// Mitsubishi GX Works2 project: B_v6_d23   PLC: Q03UDE

PROGRAM COMMON
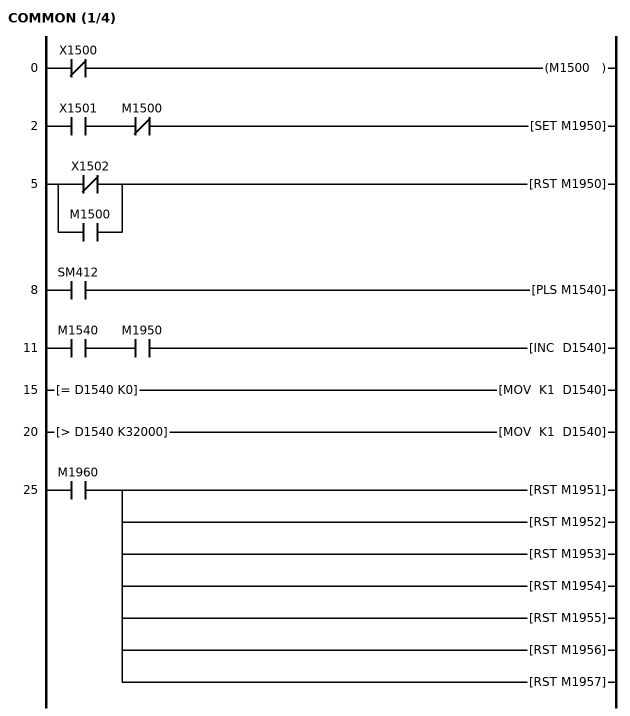
0     LDI     X1500
      OUT     M1500
2     LD      X1501
      ANI     M1500
      SET     M1950
5     LDI     X1502
      OR      M1500
      RST     M1950
8     LD      SM412
      PLS     M1540
11    LD      M1540
      AND     M1950
      INC     D1540
15    LD=     D1540 K0
      MOV     K1 D1540
20    LD>     D1540 K32000
      MOV     K1 D1540
25    LD      M1960
      RST     M1951
      RST     M1952
      RST     M1953
      RST     M1954
      RST     M1955
      RST     M1956
      RST     M1957
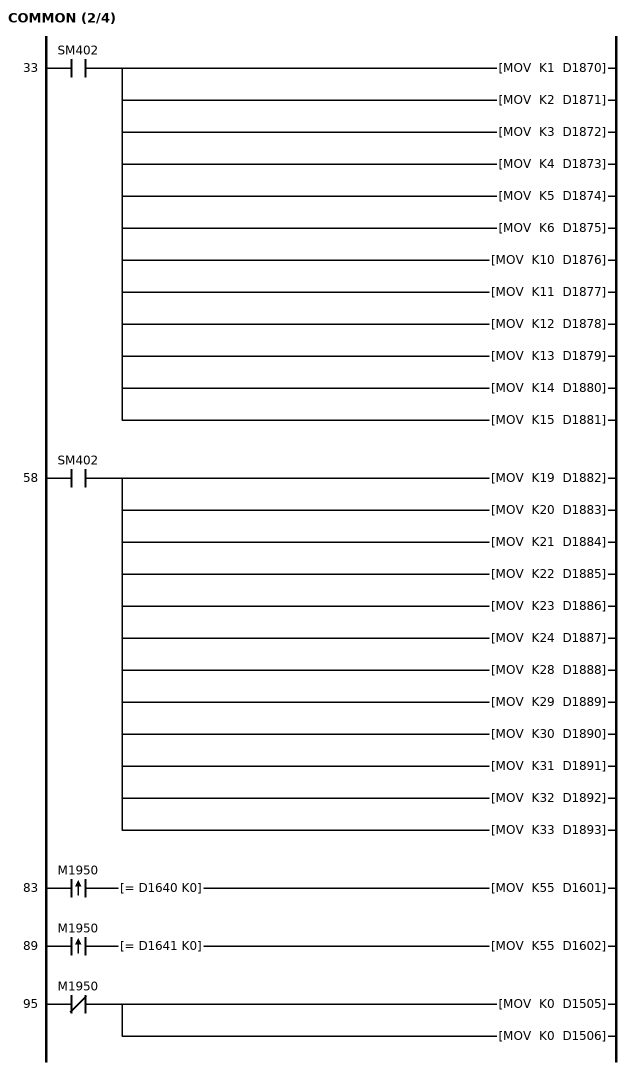
33    LD      SM402
      MOV     K1 D1870
      MOV     K2 D1871
      MOV     K3 D1872
      MOV     K4 D1873
      MOV     K5 D1874
      MOV     K6 D1875
      MOV     K10 D1876
      MOV     K11 D1877
      MOV     K12 D1878
      MOV     K13 D1879
      MOV     K14 D1880
      MOV     K15 D1881
58    LD      SM402
      MOV     K19 D1882
      MOV     K20 D1883
      MOV     K21 D1884
      MOV     K22 D1885
      MOV     K23 D1886
      MOV     K24 D1887
      MOV     K28 D1888
      MOV     K29 D1889
      MOV     K30 D1890
      MOV     K31 D1891
      MOV     K32 D1892
      MOV     K33 D1893
83    LDP     M1950
      AND=    D1640 K0
      MOV     K55 D1601
89    LDP     M1950
      AND=    D1641 K0
      MOV     K55 D1602
95    LDI     M1950
      MOV     K0 D1505
      MOV     K0 D1506
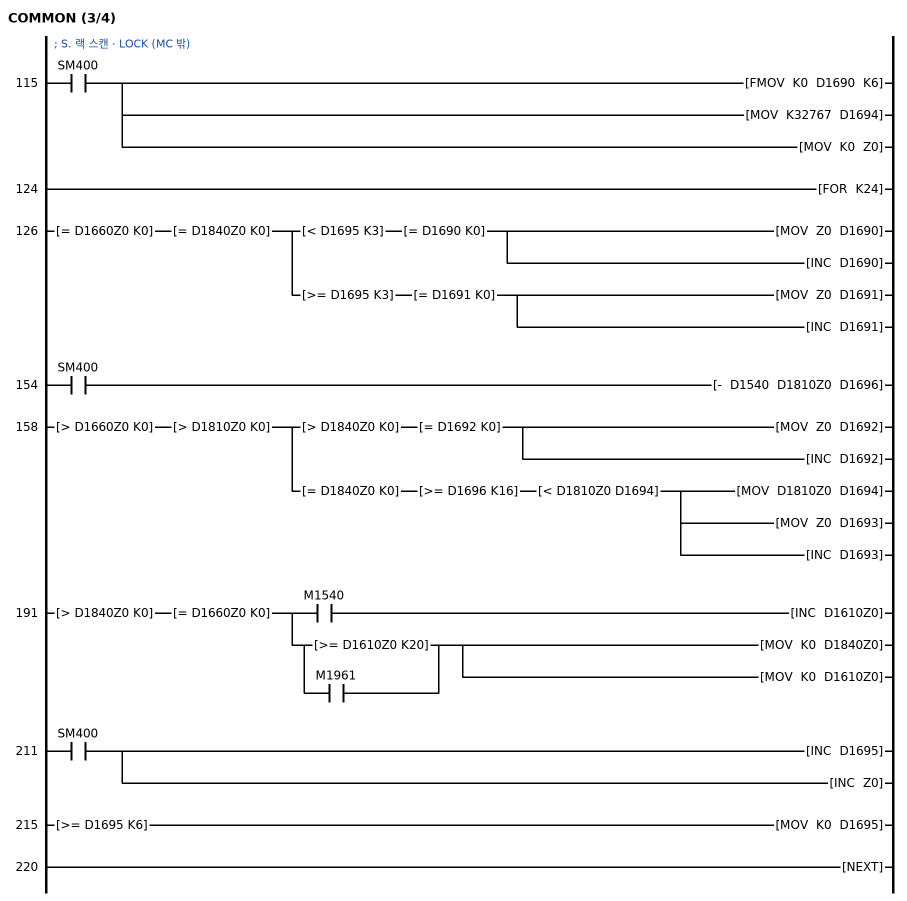
; S. 랙 스캔 · LOCK (MC 밖)
115   LD      SM400
      FMOV    K0 D1690 K6
      MOV     K32767 D1694
      MOV     K0 Z0
124   FOR     K24
126   LD=     D1660Z0 K0
      AND=    D1840Z0 K0
      MPS
      AND<    D1695 K3
      AND=    D1690 K0
      MOV     Z0 D1690
      INC     D1690
      MPP
      AND>=   D1695 K3
      AND=    D1691 K0
      MOV     Z0 D1691
      INC     D1691
154   LD      SM400
      -       D1540 D1810Z0 D1696
158   LD>     D1660Z0 K0
      AND>    D1810Z0 K0
      MPS
      AND>    D1840Z0 K0
      AND=    D1692 K0
      MOV     Z0 D1692
      INC     D1692
      MPP
      AND=    D1840Z0 K0
      AND>=   D1696 K16
      AND<    D1810Z0 D1694
      MOV     D1810Z0 D1694
      MOV     Z0 D1693
      INC     D1693
191   LD>     D1840Z0 K0
      AND=    D1660Z0 K0
      MPS
      AND     M1540
      INC     D1610Z0
      MPP
      LD>=    D1610Z0 K20
      OR      M1961
      ANB
      MOV     K0 D1840Z0
      MOV     K0 D1610Z0
211   LD      SM400
      INC     D1695
      INC     Z0
215   LD>=    D1695 K6
      MOV     K0 D1695
220   NEXT
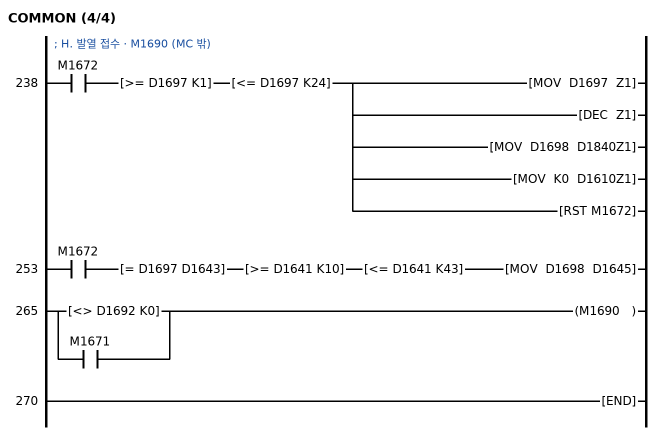
; H. 발열 접수 · M1690 (MC 밖)
238   LD      M1672
      AND>=   D1697 K1
      AND<=   D1697 K24
      MOV     D1697 Z1
      DEC     Z1
      MOV     D1698 D1840Z1
      MOV     K0 D1610Z1
      RST     M1672
253   LD      M1672
      AND=    D1697 D1643
      AND>=   D1641 K10
      AND<=   D1641 K43
      MOV     D1698 D1645
265   LD<>    D1692 K0
      OR      M1671
      OUT     M1690
270   END
END_PROGRAM

PROGRAM RFID
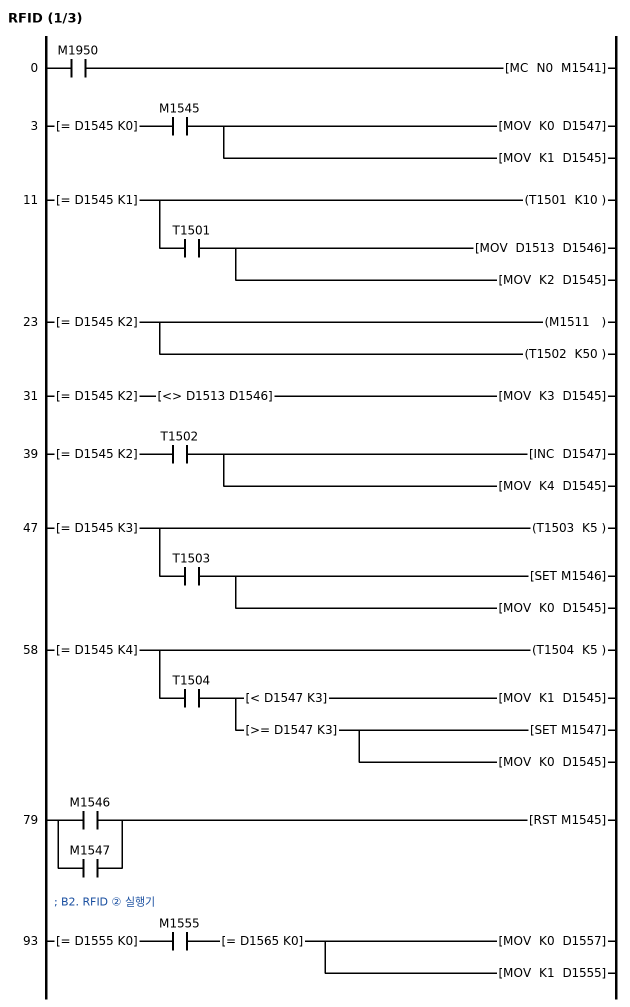
0     LD      M1950
      MC      N0 M1541
3     LD=     D1545 K0
      AND     M1545
      MOV     K0 D1547
      MOV     K1 D1545
11    LD=     D1545 K1
      OUT     T1501 K10
      AND     T1501
      MOV     D1513 D1546
      MOV     K2 D1545
23    LD=     D1545 K2
      OUT     M1511
      OUT     T1502 K50
31    LD=     D1545 K2
      AND<>   D1513 D1546
      MOV     K3 D1545
39    LD=     D1545 K2
      AND     T1502
      INC     D1547
      MOV     K4 D1545
47    LD=     D1545 K3
      OUT     T1503 K5
      AND     T1503
      SET     M1546
      MOV     K0 D1545
58    LD=     D1545 K4
      OUT     T1504 K5
      AND     T1504
      MPS
      AND<    D1547 K3
      MOV     K1 D1545
      MPP
      AND>=   D1547 K3
      SET     M1547
      MOV     K0 D1545
79    LD      M1546
      OR      M1547
      RST     M1545
; B2. RFID ② 실행기
93    LD=     D1555 K0
      AND     M1555
      AND=    D1565 K0
      MOV     K0 D1557
      MOV     K1 D1555
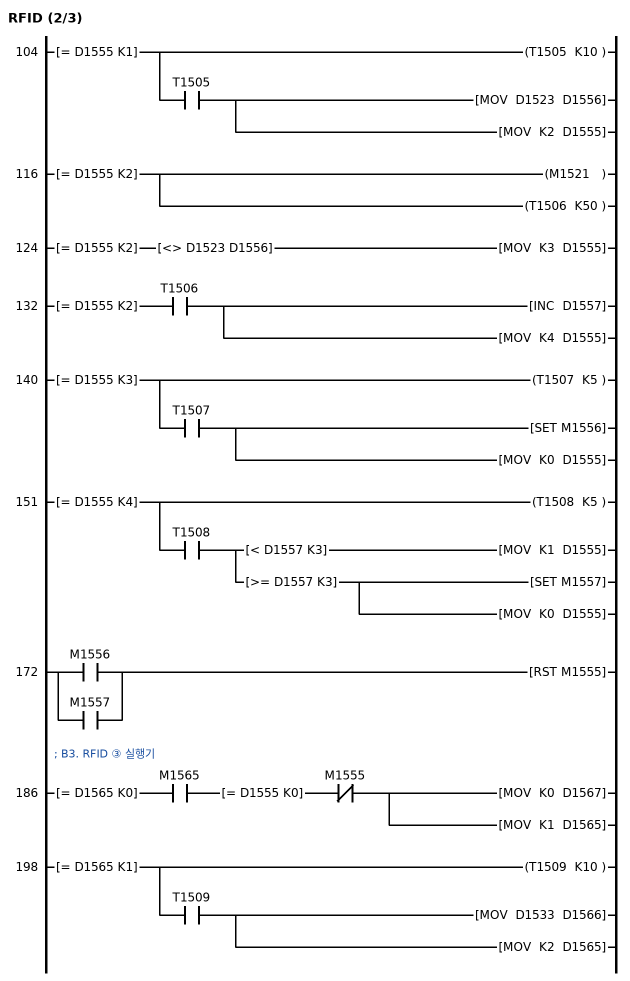
104   LD=     D1555 K1
      OUT     T1505 K10
      AND     T1505
      MOV     D1523 D1556
      MOV     K2 D1555
116   LD=     D1555 K2
      OUT     M1521
      OUT     T1506 K50
124   LD=     D1555 K2
      AND<>   D1523 D1556
      MOV     K3 D1555
132   LD=     D1555 K2
      AND     T1506
      INC     D1557
      MOV     K4 D1555
140   LD=     D1555 K3
      OUT     T1507 K5
      AND     T1507
      SET     M1556
      MOV     K0 D1555
151   LD=     D1555 K4
      OUT     T1508 K5
      AND     T1508
      MPS
      AND<    D1557 K3
      MOV     K1 D1555
      MPP
      AND>=   D1557 K3
      SET     M1557
      MOV     K0 D1555
172   LD      M1556
      OR      M1557
      RST     M1555
; B3. RFID ③ 실행기
186   LD=     D1565 K0
      AND     M1565
      AND=    D1555 K0
      ANI     M1555
      MOV     K0 D1567
      MOV     K1 D1565
198   LD=     D1565 K1
      OUT     T1509 K10
      AND     T1509
      MOV     D1533 D1566
      MOV     K2 D1565
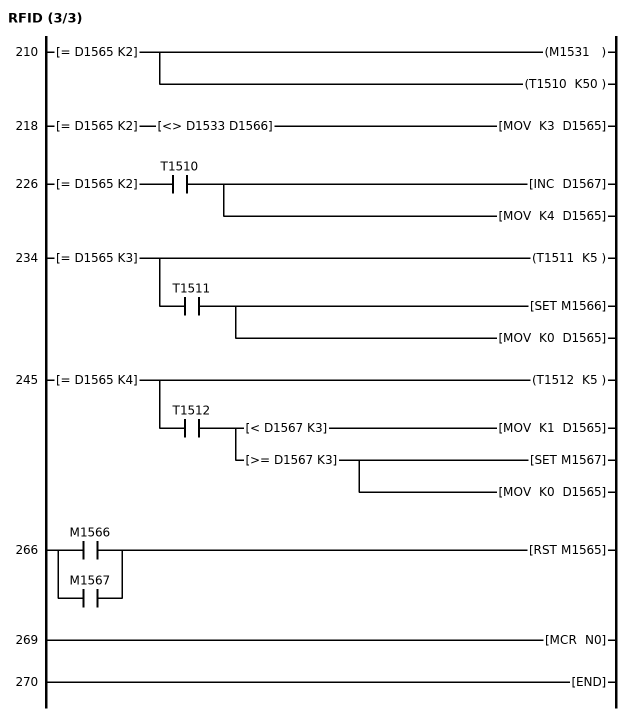
210   LD=     D1565 K2
      OUT     M1531
      OUT     T1510 K50
218   LD=     D1565 K2
      AND<>   D1533 D1566
      MOV     K3 D1565
226   LD=     D1565 K2
      AND     T1510
      INC     D1567
      MOV     K4 D1565
234   LD=     D1565 K3
      OUT     T1511 K5
      AND     T1511
      SET     M1566
      MOV     K0 D1565
245   LD=     D1565 K4
      OUT     T1512 K5
      AND     T1512
      MPS
      AND<    D1567 K3
      MOV     K1 D1565
      MPP
      AND>=   D1567 K3
      SET     M1567
      MOV     K0 D1565
266   LD      M1566
      OR      M1567
      RST     M1565
269   MCR     N0
270   END
END_PROGRAM

PROGRAM INFEED
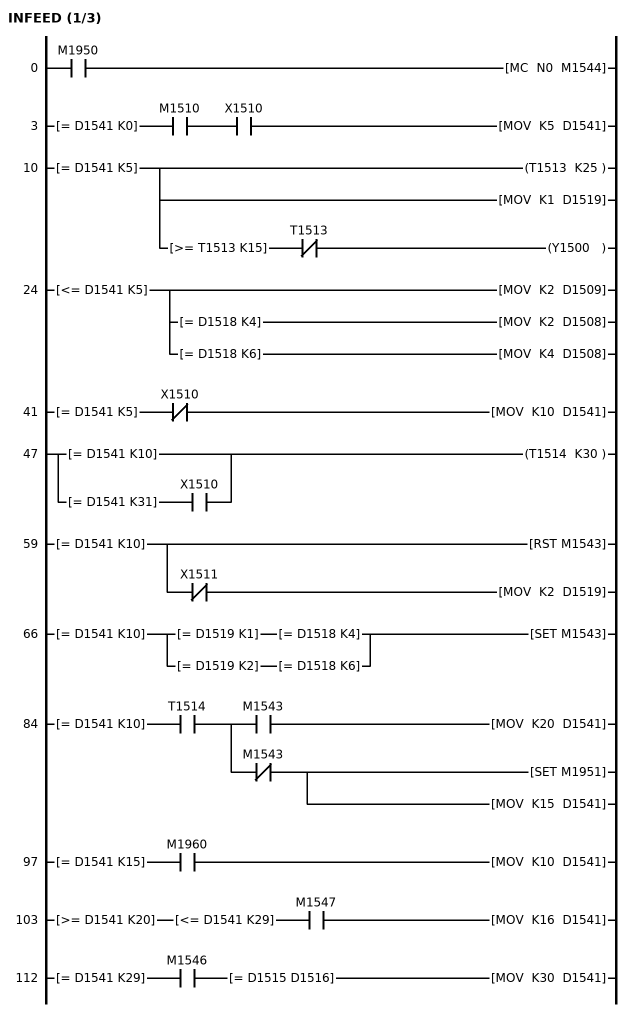
0     LD      M1950
      MC      N0 M1544
3     LD=     D1541 K0
      AND     M1510
      AND     X1510
      MOV     K5 D1541
10    LD=     D1541 K5
      OUT     T1513 K25
      MOV     K1 D1519
      AND>=   T1513 K15
      ANI     T1513
      OUT     Y1500
24    LD<=    D1541 K5
      MOV     K2 D1509
      MPS
      AND=    D1518 K4
      MOV     K2 D1508
      MPP
      AND=    D1518 K6
      MOV     K4 D1508
41    LD=     D1541 K5
      ANI     X1510
      MOV     K10 D1541
47    LD=     D1541 K10
      LD=     D1541 K31
      AND     X1510
      ORB
      OUT     T1514 K30
59    LD=     D1541 K10
      RST     M1543
      ANI     X1511
      MOV     K2 D1519
66    LD=     D1541 K10
      LD=     D1519 K1
      AND=    D1518 K4
      LD=     D1519 K2
      AND=    D1518 K6
      ORB
      ANB
      SET     M1543
84    LD=     D1541 K10
      AND     T1514
      MPS
      AND     M1543
      MOV     K20 D1541
      MPP
      ANI     M1543
      SET     M1951
      MOV     K15 D1541
97    LD=     D1541 K15
      AND     M1960
      MOV     K10 D1541
103   LD>=    D1541 K20
      AND<=   D1541 K29
      AND     M1547
      MOV     K16 D1541
112   LD=     D1541 K29
      AND     M1546
      AND=    D1515 D1516
      MOV     K30 D1541
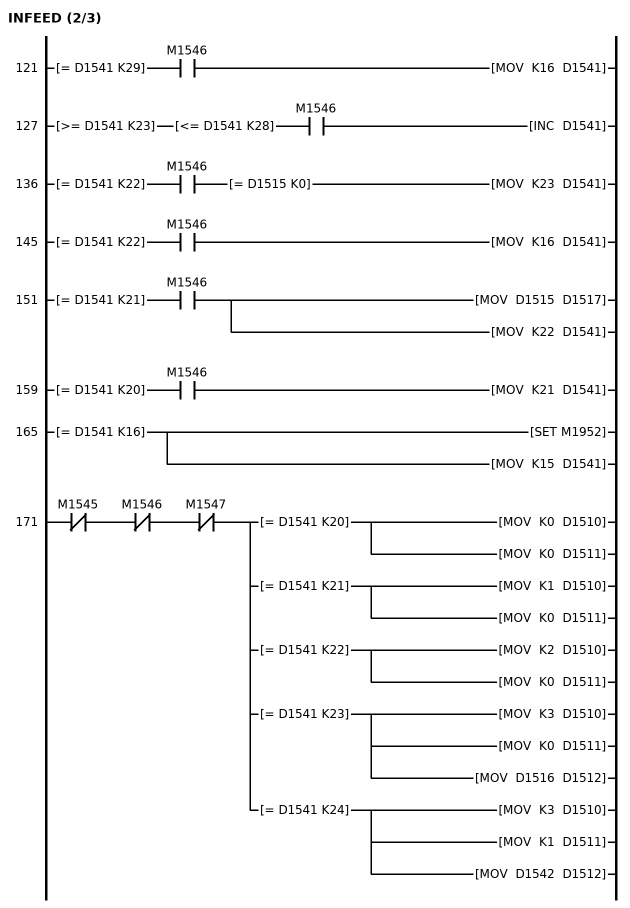
121   LD=     D1541 K29
      AND     M1546
      MOV     K16 D1541
127   LD>=    D1541 K23
      AND<=   D1541 K28
      AND     M1546
      INC     D1541
136   LD=     D1541 K22
      AND     M1546
      AND=    D1515 K0
      MOV     K23 D1541
145   LD=     D1541 K22
      AND     M1546
      MOV     K16 D1541
151   LD=     D1541 K21
      AND     M1546
      MOV     D1515 D1517
      MOV     K22 D1541
159   LD=     D1541 K20
      AND     M1546
      MOV     K21 D1541
165   LD=     D1541 K16
      SET     M1952
      MOV     K15 D1541
171   LDI     M1545
      ANI     M1546
      ANI     M1547
      MPS
      AND=    D1541 K20
      MOV     K0 D1510
      MOV     K0 D1511
      MRD
      AND=    D1541 K21
      MOV     K1 D1510
      MOV     K0 D1511
      MRD
      AND=    D1541 K22
      MOV     K2 D1510
      MOV     K0 D1511
      MRD
      AND=    D1541 K23
      MOV     K3 D1510
      MOV     K0 D1511
      MOV     D1516 D1512
      MPP
      AND=    D1541 K24
      MOV     K3 D1510
      MOV     K1 D1511
      MOV     D1542 D1512
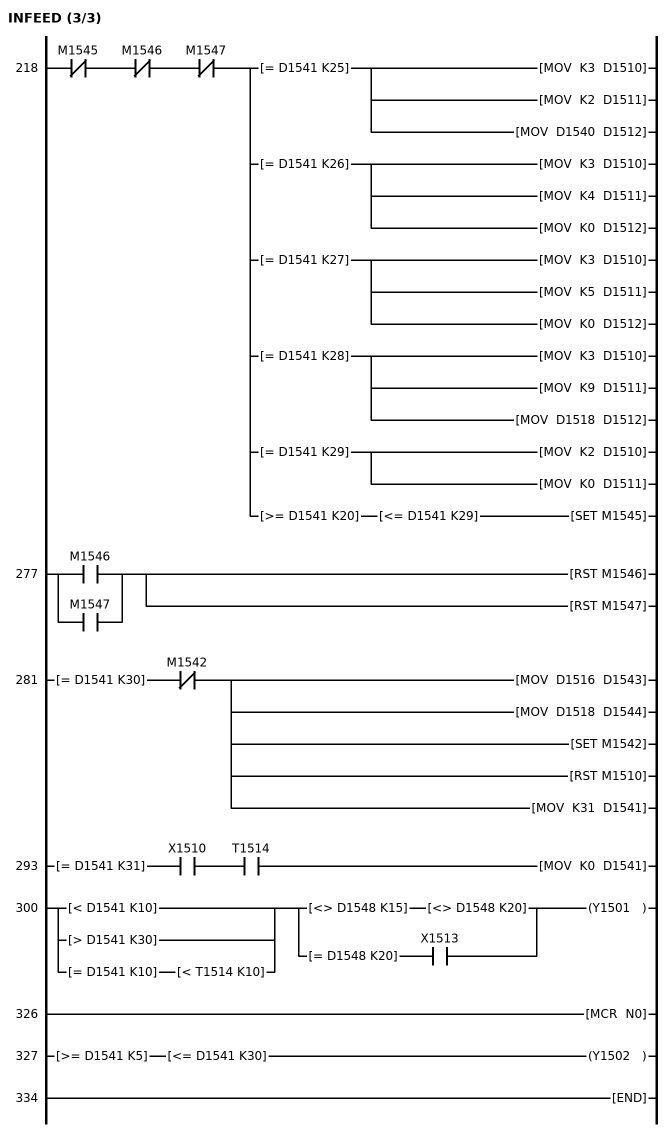
218   LDI     M1545
      ANI     M1546
      ANI     M1547
      MPS
      AND=    D1541 K25
      MOV     K3 D1510
      MOV     K2 D1511
      MOV     D1540 D1512
      MRD
      AND=    D1541 K26
      MOV     K3 D1510
      MOV     K4 D1511
      MOV     K0 D1512
      MRD
      AND=    D1541 K27
      MOV     K3 D1510
      MOV     K5 D1511
      MOV     K0 D1512
      MRD
      AND=    D1541 K28
      MOV     K3 D1510
      MOV     K9 D1511
      MOV     D1518 D1512
      MRD
      AND=    D1541 K29
      MOV     K2 D1510
      MOV     K0 D1511
      MPP
      AND>=   D1541 K20
      AND<=   D1541 K29
      SET     M1545
277   LD      M1546
      OR      M1547
      RST     M1546
      RST     M1547
281   LD=     D1541 K30
      ANI     M1542
      MOV     D1516 D1543
      MOV     D1518 D1544
      SET     M1542
      RST     M1510
      MOV     K31 D1541
293   LD=     D1541 K31
      AND     X1510
      AND     T1514
      MOV     K0 D1541
300   LD<     D1541 K10
      OR>     D1541 K30
      LD=     D1541 K10
      AND<    T1514 K10
      ORB
      LD<>    D1548 K15
      AND<>   D1548 K20
      LD=     D1548 K20
      AND     X1513
      ORB
      ANB
      OUT     Y1501
326   MCR     N0
327   LD>=    D1541 K5
      AND<=   D1541 K30
      OUT     Y1502
334   END
END_PROGRAM

PROGRAM CRANE
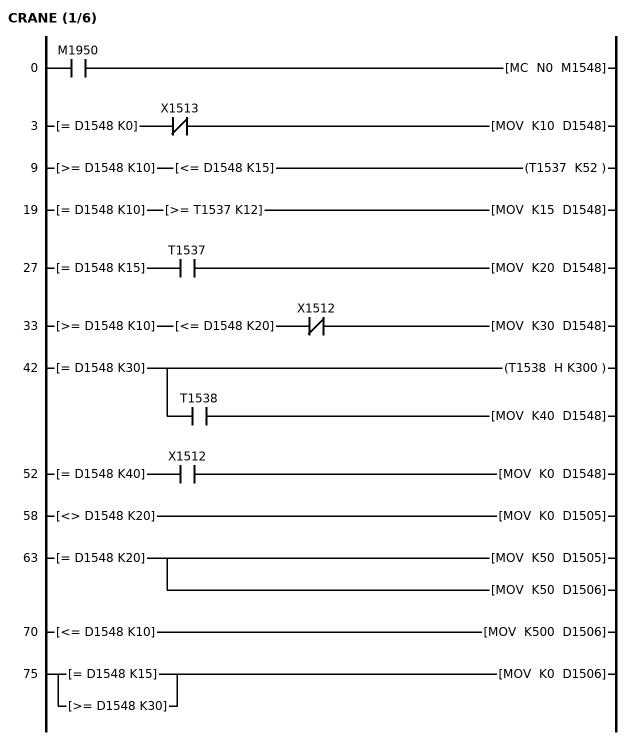
0     LD      M1950
      MC      N0 M1548
3     LD=     D1548 K0
      ANI     X1513
      MOV     K10 D1548
9     LD>=    D1548 K10
      AND<=   D1548 K15
      OUT     T1537 K52
19    LD=     D1548 K10
      AND>=   T1537 K12
      MOV     K15 D1548
27    LD=     D1548 K15
      AND     T1537
      MOV     K20 D1548
33    LD>=    D1548 K10
      AND<=   D1548 K20
      ANI     X1512
      MOV     K30 D1548
42    LD=     D1548 K30
      OUTH    T1538 K300
      AND     T1538
      MOV     K40 D1548
52    LD=     D1548 K40
      AND     X1512
      MOV     K0 D1548
58    LD<>    D1548 K20
      MOV     K0 D1505
63    LD=     D1548 K20
      MOV     K50 D1505
      MOV     K50 D1506
70    LD<=    D1548 K10
      MOV     K500 D1506
75    LD=     D1548 K15
      OR>=    D1548 K30
      MOV     K0 D1506
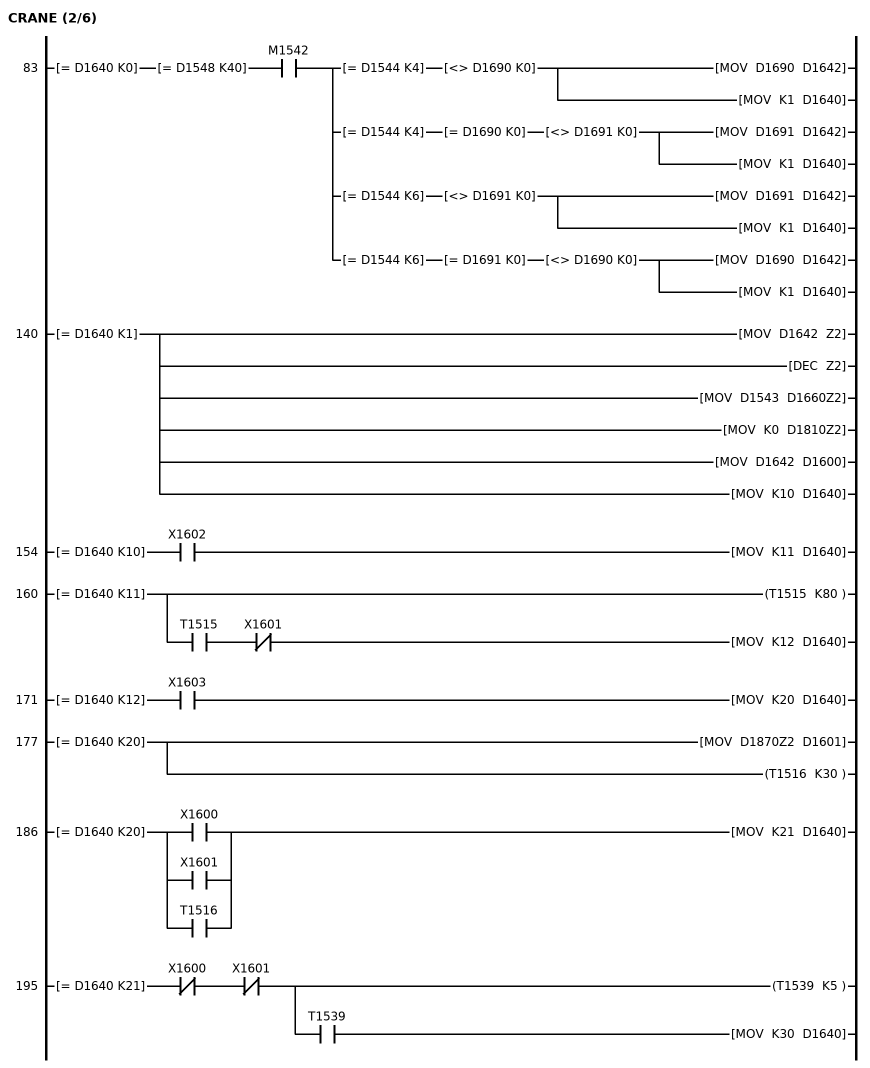
83    LD=     D1640 K0
      AND=    D1548 K40
      AND     M1542
      MPS
      AND=    D1544 K4
      AND<>   D1690 K0
      MOV     D1690 D1642
      MOV     K1 D1640
      MRD
      AND=    D1544 K4
      AND=    D1690 K0
      AND<>   D1691 K0
      MOV     D1691 D1642
      MOV     K1 D1640
      MRD
      AND=    D1544 K6
      AND<>   D1691 K0
      MOV     D1691 D1642
      MOV     K1 D1640
      MPP
      AND=    D1544 K6
      AND=    D1691 K0
      AND<>   D1690 K0
      MOV     D1690 D1642
      MOV     K1 D1640
140   LD=     D1640 K1
      MOV     D1642 Z2
      DEC     Z2
      MOV     D1543 D1660Z2
      MOV     K0 D1810Z2
      MOV     D1642 D1600
      MOV     K10 D1640
154   LD=     D1640 K10
      AND     X1602
      MOV     K11 D1640
160   LD=     D1640 K11
      OUT     T1515 K80
      AND     T1515
      ANI     X1601
      MOV     K12 D1640
171   LD=     D1640 K12
      AND     X1603
      MOV     K20 D1640
177   LD=     D1640 K20
      MOV     D1870Z2 D1601
      OUT     T1516 K30
186   LD=     D1640 K20
      LD      X1600
      OR      X1601
      OR      T1516
      ANB
      MOV     K21 D1640
195   LD=     D1640 K21
      ANI     X1600
      ANI     X1601
      OUT     T1539 K5
      AND     T1539
      MOV     K30 D1640
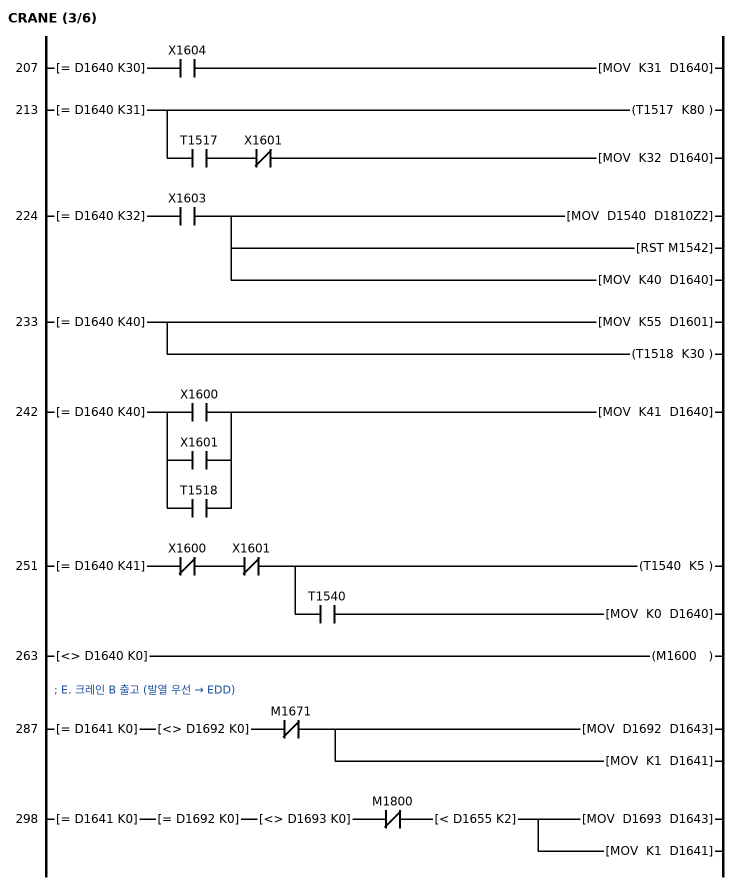
207   LD=     D1640 K30
      AND     X1604
      MOV     K31 D1640
213   LD=     D1640 K31
      OUT     T1517 K80
      AND     T1517
      ANI     X1601
      MOV     K32 D1640
224   LD=     D1640 K32
      AND     X1603
      MOV     D1540 D1810Z2
      RST     M1542
      MOV     K40 D1640
233   LD=     D1640 K40
      MOV     K55 D1601
      OUT     T1518 K30
242   LD=     D1640 K40
      LD      X1600
      OR      X1601
      OR      T1518
      ANB
      MOV     K41 D1640
251   LD=     D1640 K41
      ANI     X1600
      ANI     X1601
      OUT     T1540 K5
      AND     T1540
      MOV     K0 D1640
263   LD<>    D1640 K0
      OUT     M1600
; E. 크레인 B 출고 (발열 우선 → EDD)
287   LD=     D1641 K0
      AND<>   D1692 K0
      ANI     M1671
      MOV     D1692 D1643
      MOV     K1 D1641
298   LD=     D1641 K0
      AND=    D1692 K0
      AND<>   D1693 K0
      ANI     M1800
      AND<    D1655 K2
      MOV     D1693 D1643
      MOV     K1 D1641
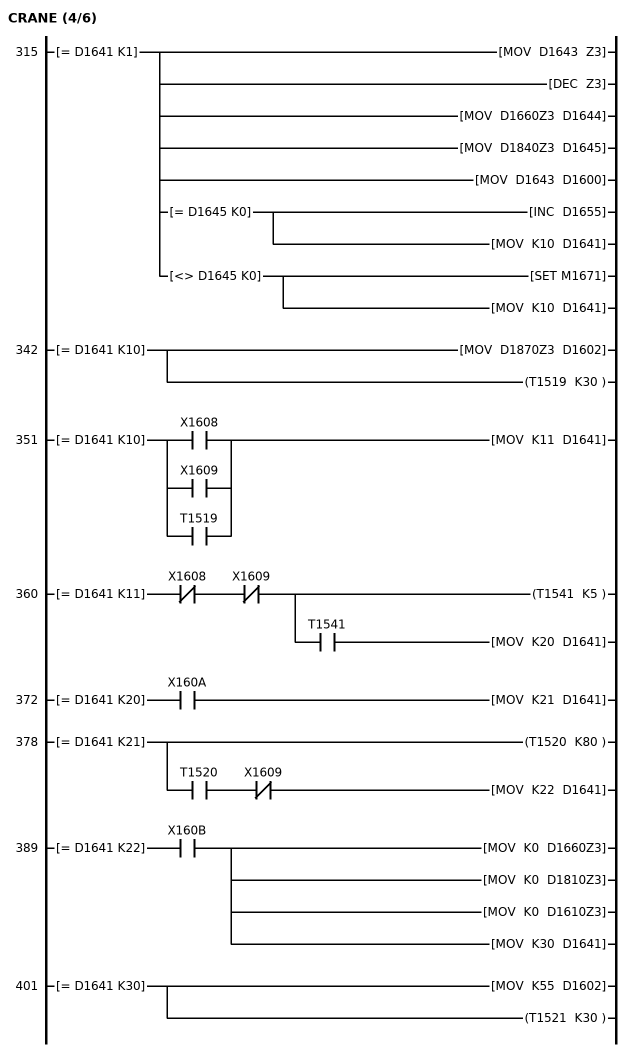
315   LD=     D1641 K1
      MOV     D1643 Z3
      DEC     Z3
      MOV     D1660Z3 D1644
      MOV     D1840Z3 D1645
      MOV     D1643 D1600
      MPS
      AND=    D1645 K0
      INC     D1655
      MOV     K10 D1641
      MPP
      AND<>   D1645 K0
      SET     M1671
      MOV     K10 D1641
342   LD=     D1641 K10
      MOV     D1870Z3 D1602
      OUT     T1519 K30
351   LD=     D1641 K10
      LD      X1608
      OR      X1609
      OR      T1519
      ANB
      MOV     K11 D1641
360   LD=     D1641 K11
      ANI     X1608
      ANI     X1609
      OUT     T1541 K5
      AND     T1541
      MOV     K20 D1641
372   LD=     D1641 K20
      AND     X160A
      MOV     K21 D1641
378   LD=     D1641 K21
      OUT     T1520 K80
      AND     T1520
      ANI     X1609
      MOV     K22 D1641
389   LD=     D1641 K22
      AND     X160B
      MOV     K0 D1660Z3
      MOV     K0 D1810Z3
      MOV     K0 D1610Z3
      MOV     K30 D1641
401   LD=     D1641 K30
      MOV     K55 D1602
      OUT     T1521 K30
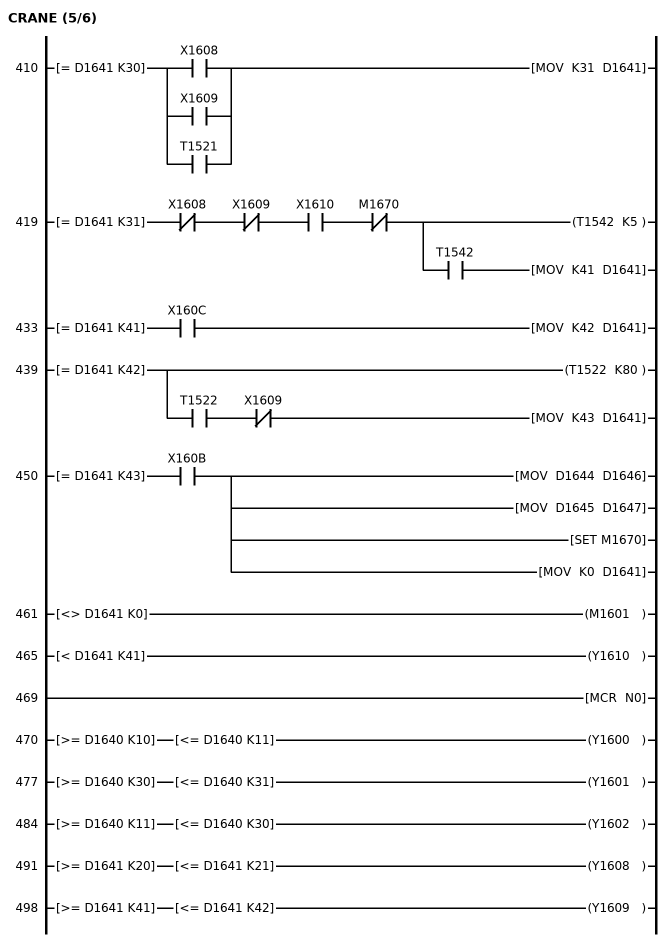
410   LD=     D1641 K30
      LD      X1608
      OR      X1609
      OR      T1521
      ANB
      MOV     K31 D1641
419   LD=     D1641 K31
      ANI     X1608
      ANI     X1609
      AND     X1610
      ANI     M1670
      OUT     T1542 K5
      AND     T1542
      MOV     K41 D1641
433   LD=     D1641 K41
      AND     X160C
      MOV     K42 D1641
439   LD=     D1641 K42
      OUT     T1522 K80
      AND     T1522
      ANI     X1609
      MOV     K43 D1641
450   LD=     D1641 K43
      AND     X160B
      MOV     D1644 D1646
      MOV     D1645 D1647
      SET     M1670
      MOV     K0 D1641
461   LD<>    D1641 K0
      OUT     M1601
465   LD<     D1641 K41
      OUT     Y1610
469   MCR     N0
470   LD>=    D1640 K10
      AND<=   D1640 K11
      OUT     Y1600
477   LD>=    D1640 K30
      AND<=   D1640 K31
      OUT     Y1601
484   LD>=    D1640 K11
      AND<=   D1640 K30
      OUT     Y1602
491   LD>=    D1641 K20
      AND<=   D1641 K21
      OUT     Y1608
498   LD>=    D1641 K41
      AND<=   D1641 K42
      OUT     Y1609
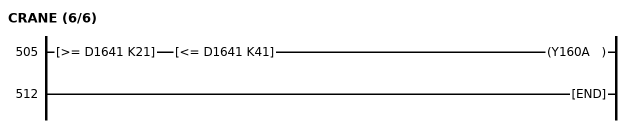
505   LD>=    D1641 K21
      AND<=   D1641 K41
      OUT     Y160A
512   END
END_PROGRAM

PROGRAM SORT1
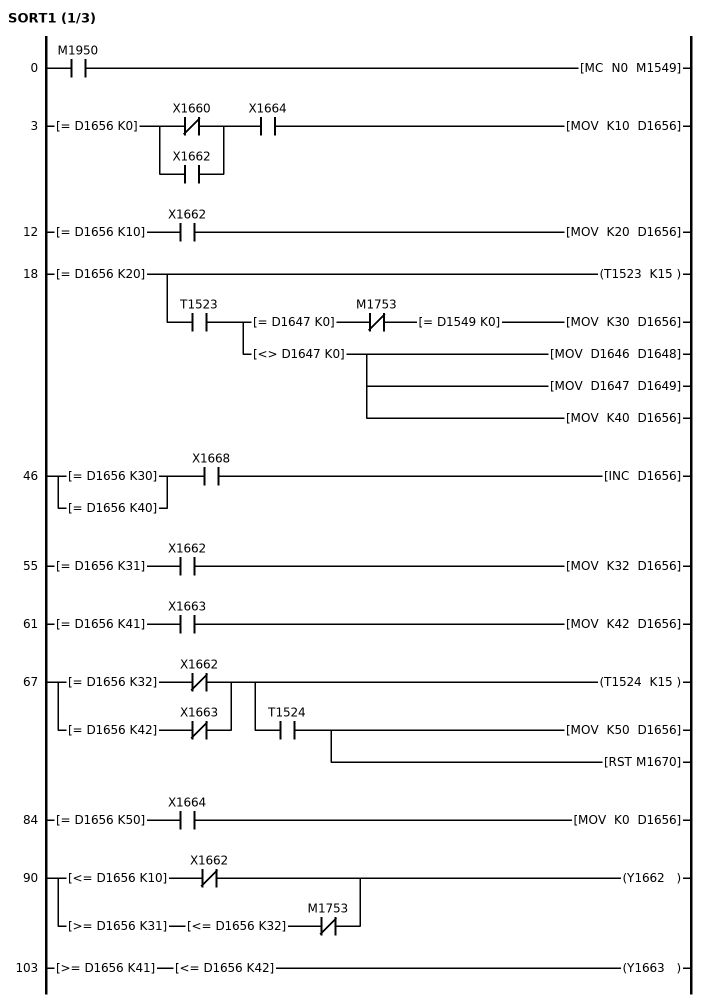
0     LD      M1950
      MC      N0 M1549
3     LD=     D1656 K0
      LDI     X1660
      OR      X1662
      ANB
      AND     X1664
      MOV     K10 D1656
12    LD=     D1656 K10
      AND     X1662
      MOV     K20 D1656
18    LD=     D1656 K20
      OUT     T1523 K15
      AND     T1523
      MPS
      AND=    D1647 K0
      ANI     M1753
      AND=    D1549 K0
      MOV     K30 D1656
      MPP
      AND<>   D1647 K0
      MOV     D1646 D1648
      MOV     D1647 D1649
      MOV     K40 D1656
46    LD=     D1656 K30
      OR=     D1656 K40
      AND     X1668
      INC     D1656
55    LD=     D1656 K31
      AND     X1662
      MOV     K32 D1656
61    LD=     D1656 K41
      AND     X1663
      MOV     K42 D1656
67    LD=     D1656 K32
      ANI     X1662
      LD=     D1656 K42
      ANI     X1663
      ORB
      OUT     T1524 K15
      AND     T1524
      MOV     K50 D1656
      RST     M1670
84    LD=     D1656 K50
      AND     X1664
      MOV     K0 D1656
90    LD<=    D1656 K10
      ANI     X1662
      LD>=    D1656 K31
      AND<=   D1656 K32
      ANI     M1753
      ORB
      OUT     Y1662
103   LD>=    D1656 K41
      AND<=   D1656 K42
      OUT     Y1663
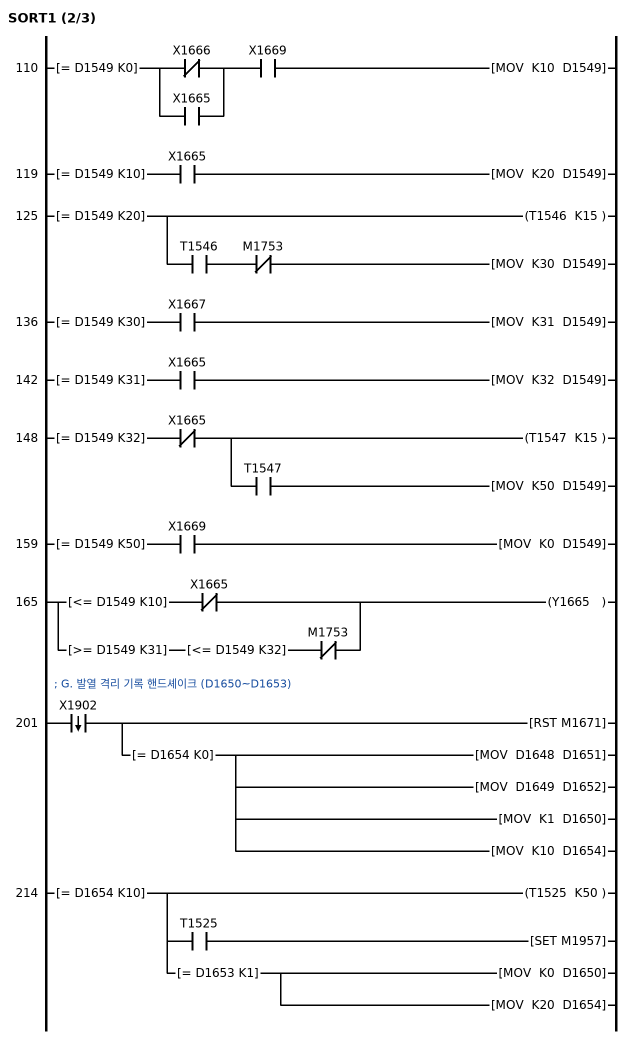
110   LD=     D1549 K0
      LDI     X1666
      OR      X1665
      ANB
      AND     X1669
      MOV     K10 D1549
119   LD=     D1549 K10
      AND     X1665
      MOV     K20 D1549
125   LD=     D1549 K20
      OUT     T1546 K15
      AND     T1546
      ANI     M1753
      MOV     K30 D1549
136   LD=     D1549 K30
      AND     X1667
      MOV     K31 D1549
142   LD=     D1549 K31
      AND     X1665
      MOV     K32 D1549
148   LD=     D1549 K32
      ANI     X1665
      OUT     T1547 K15
      AND     T1547
      MOV     K50 D1549
159   LD=     D1549 K50
      AND     X1669
      MOV     K0 D1549
165   LD<=    D1549 K10
      ANI     X1665
      LD>=    D1549 K31
      AND<=   D1549 K32
      ANI     M1753
      ORB
      OUT     Y1665
; G. 발열 격리 기록 핸드셰이크 (D1650~D1653)
201   LDF     X1902
      RST     M1671
      AND=    D1654 K0
      MOV     D1648 D1651
      MOV     D1649 D1652
      MOV     K1 D1650
      MOV     K10 D1654
214   LD=     D1654 K10
      OUT     T1525 K50
      MPS
      AND     T1525
      SET     M1957
      MPP
      AND=    D1653 K1
      MOV     K0 D1650
      MOV     K20 D1654
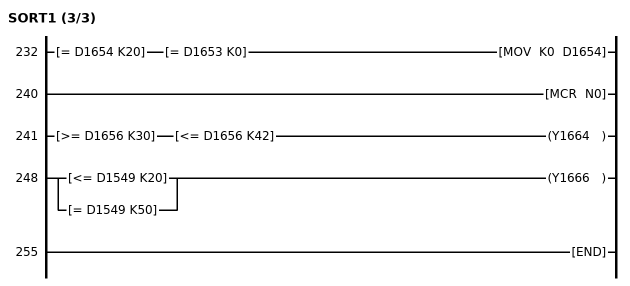
232   LD=     D1654 K20
      AND=    D1653 K0
      MOV     K0 D1654
240   MCR     N0
241   LD>=    D1656 K30
      AND<=   D1656 K42
      OUT     Y1664
248   LD<=    D1549 K20
      OR=     D1549 K50
      OUT     Y1666
255   END
END_PROGRAM

PROGRAM INSPECT
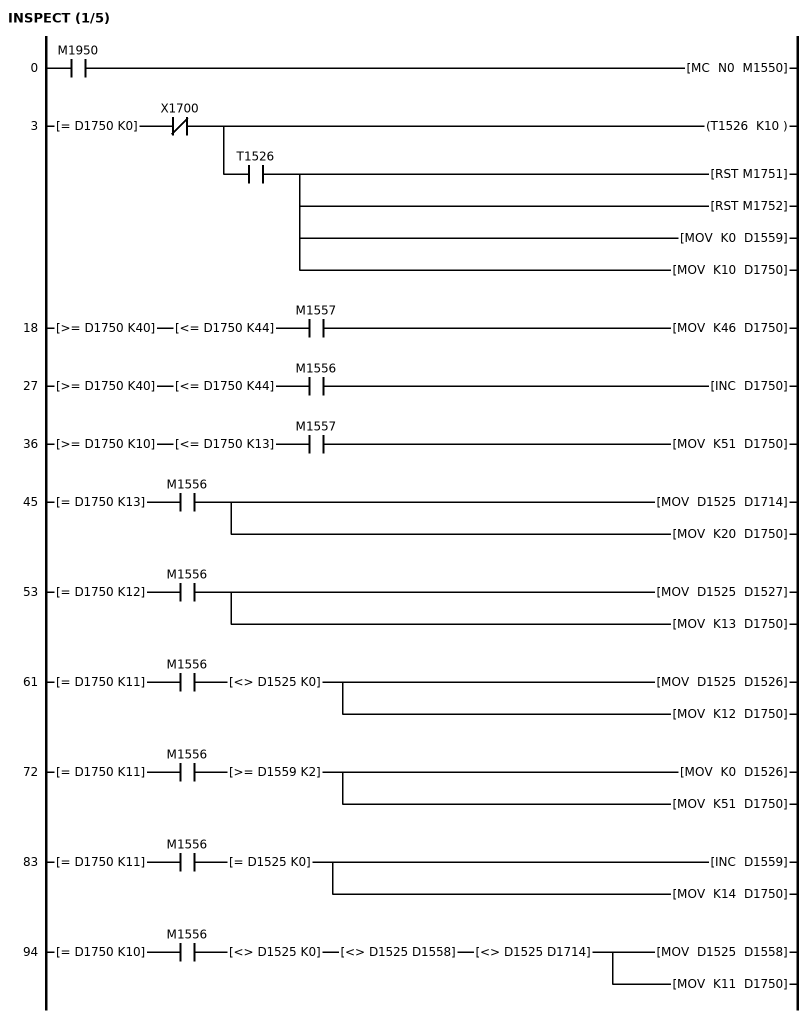
0     LD      M1950
      MC      N0 M1550
3     LD=     D1750 K0
      ANI     X1700
      OUT     T1526 K10
      AND     T1526
      RST     M1751
      RST     M1752
      MOV     K0 D1559
      MOV     K10 D1750
18    LD>=    D1750 K40
      AND<=   D1750 K44
      AND     M1557
      MOV     K46 D1750
27    LD>=    D1750 K40
      AND<=   D1750 K44
      AND     M1556
      INC     D1750
36    LD>=    D1750 K10
      AND<=   D1750 K13
      AND     M1557
      MOV     K51 D1750
45    LD=     D1750 K13
      AND     M1556
      MOV     D1525 D1714
      MOV     K20 D1750
53    LD=     D1750 K12
      AND     M1556
      MOV     D1525 D1527
      MOV     K13 D1750
61    LD=     D1750 K11
      AND     M1556
      AND<>   D1525 K0
      MOV     D1525 D1526
      MOV     K12 D1750
72    LD=     D1750 K11
      AND     M1556
      AND>=   D1559 K2
      MOV     K0 D1526
      MOV     K51 D1750
83    LD=     D1750 K11
      AND     M1556
      AND=    D1525 K0
      INC     D1559
      MOV     K14 D1750
94    LD=     D1750 K10
      AND     M1556
      AND<>   D1525 K0
      AND<>   D1525 D1558
      AND<>   D1525 D1714
      MOV     D1525 D1558
      MOV     K11 D1750
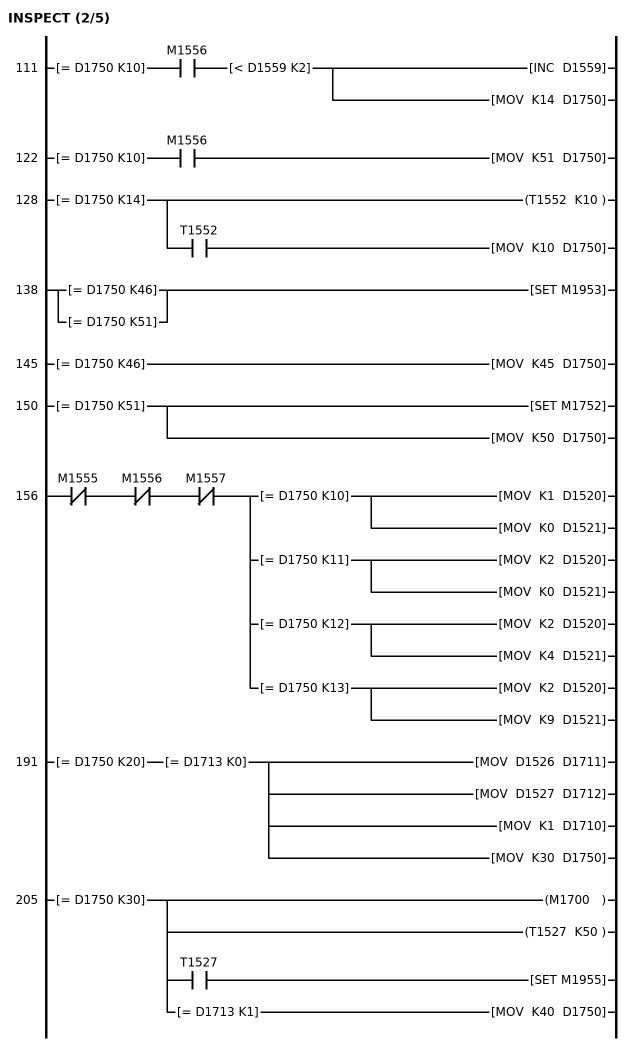
111   LD=     D1750 K10
      AND     M1556
      AND<    D1559 K2
      INC     D1559
      MOV     K14 D1750
122   LD=     D1750 K10
      AND     M1556
      MOV     K51 D1750
128   LD=     D1750 K14
      OUT     T1552 K10
      AND     T1552
      MOV     K10 D1750
138   LD=     D1750 K46
      OR=     D1750 K51
      SET     M1953
145   LD=     D1750 K46
      MOV     K45 D1750
150   LD=     D1750 K51
      SET     M1752
      MOV     K50 D1750
156   LDI     M1555
      ANI     M1556
      ANI     M1557
      MPS
      AND=    D1750 K10
      MOV     K1 D1520
      MOV     K0 D1521
      MRD
      AND=    D1750 K11
      MOV     K2 D1520
      MOV     K0 D1521
      MRD
      AND=    D1750 K12
      MOV     K2 D1520
      MOV     K4 D1521
      MPP
      AND=    D1750 K13
      MOV     K2 D1520
      MOV     K9 D1521
191   LD=     D1750 K20
      AND=    D1713 K0
      MOV     D1526 D1711
      MOV     D1527 D1712
      MOV     K1 D1710
      MOV     K30 D1750
205   LD=     D1750 K30
      OUT     M1700
      OUT     T1527 K50
      MPS
      AND     T1527
      SET     M1955
      MPP
      AND=    D1713 K1
      MOV     K40 D1750
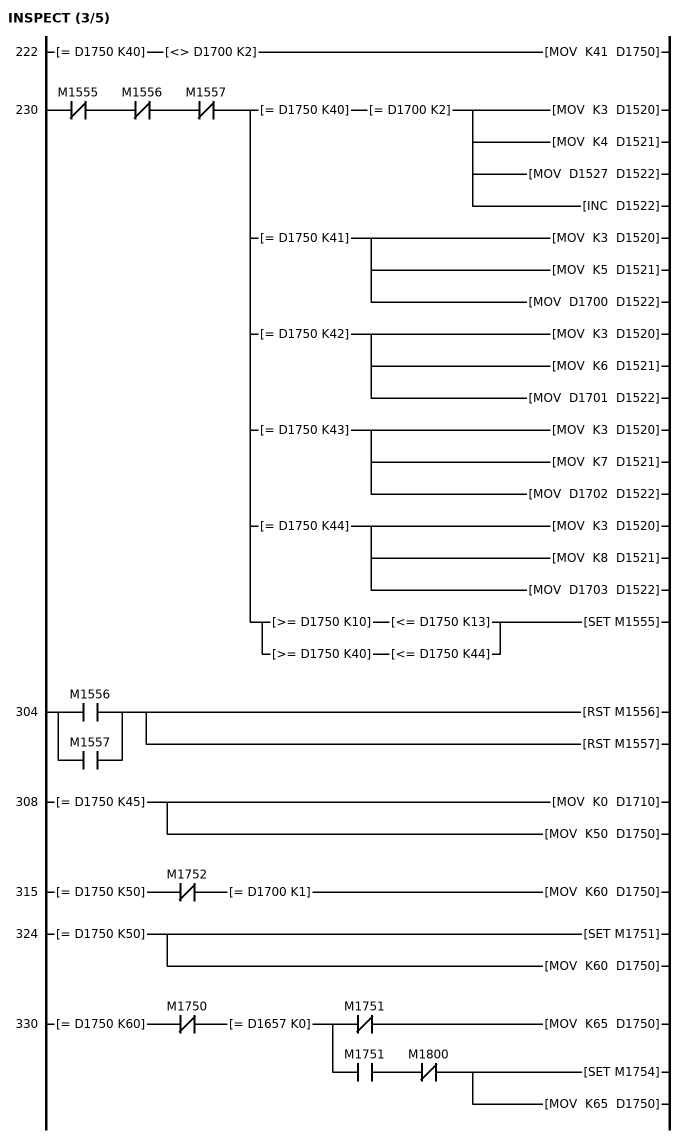
222   LD=     D1750 K40
      AND<>   D1700 K2
      MOV     K41 D1750
230   LDI     M1555
      ANI     M1556
      ANI     M1557
      MPS
      AND=    D1750 K40
      AND=    D1700 K2
      MOV     K3 D1520
      MOV     K4 D1521
      MOV     D1527 D1522
      INC     D1522
      MRD
      AND=    D1750 K41
      MOV     K3 D1520
      MOV     K5 D1521
      MOV     D1700 D1522
      MRD
      AND=    D1750 K42
      MOV     K3 D1520
      MOV     K6 D1521
      MOV     D1701 D1522
      MRD
      AND=    D1750 K43
      MOV     K3 D1520
      MOV     K7 D1521
      MOV     D1702 D1522
      MRD
      AND=    D1750 K44
      MOV     K3 D1520
      MOV     K8 D1521
      MOV     D1703 D1522
      MPP
      LD>=    D1750 K10
      AND<=   D1750 K13
      LD>=    D1750 K40
      AND<=   D1750 K44
      ORB
      ANB
      SET     M1555
304   LD      M1556
      OR      M1557
      RST     M1556
      RST     M1557
308   LD=     D1750 K45
      MOV     K0 D1710
      MOV     K50 D1750
315   LD=     D1750 K50
      ANI     M1752
      AND=    D1700 K1
      MOV     K60 D1750
324   LD=     D1750 K50
      SET     M1751
      MOV     K60 D1750
330   LD=     D1750 K60
      ANI     M1750
      AND=    D1657 K0
      MPS
      ANI     M1751
      MOV     K65 D1750
      MPP
      AND     M1751
      ANI     M1800
      SET     M1754
      MOV     K65 D1750
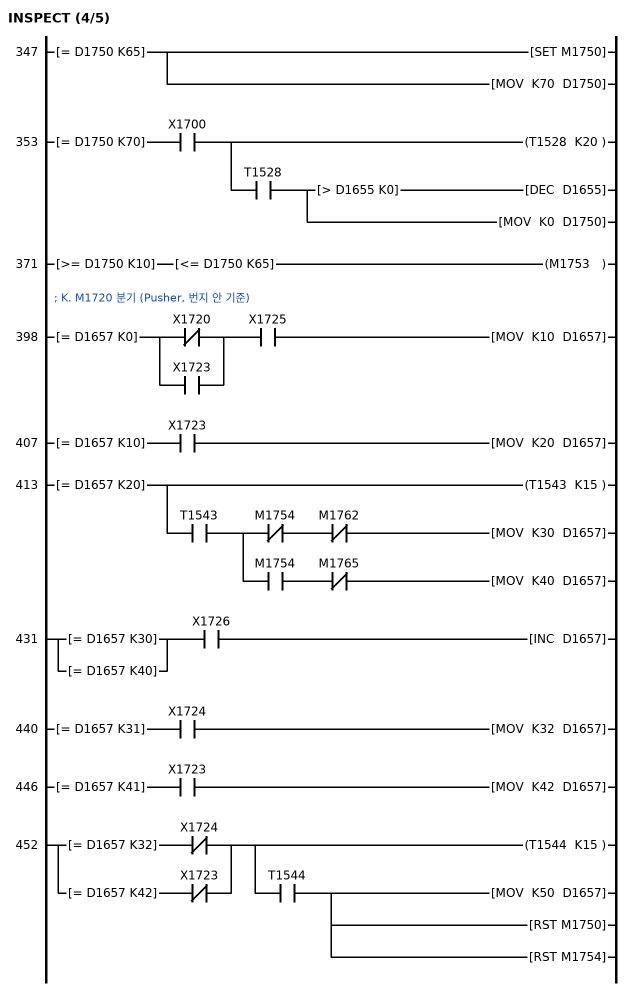
347   LD=     D1750 K65
      SET     M1750
      MOV     K70 D1750
353   LD=     D1750 K70
      AND     X1700
      OUT     T1528 K20
      AND     T1528
      MPS
      AND>    D1655 K0
      DEC     D1655
      MPP
      MOV     K0 D1750
371   LD>=    D1750 K10
      AND<=   D1750 K65
      OUT     M1753
; K. M1720 분기 (Pusher, 번지 안 기준)
398   LD=     D1657 K0
      LDI     X1720
      OR      X1723
      ANB
      AND     X1725
      MOV     K10 D1657
407   LD=     D1657 K10
      AND     X1723
      MOV     K20 D1657
413   LD=     D1657 K20
      OUT     T1543 K15
      AND     T1543
      MPS
      ANI     M1754
      ANI     M1762
      MOV     K30 D1657
      MPP
      AND     M1754
      ANI     M1765
      MOV     K40 D1657
431   LD=     D1657 K30
      OR=     D1657 K40
      AND     X1726
      INC     D1657
440   LD=     D1657 K31
      AND     X1724
      MOV     K32 D1657
446   LD=     D1657 K41
      AND     X1723
      MOV     K42 D1657
452   LD=     D1657 K32
      ANI     X1724
      LD=     D1657 K42
      ANI     X1723
      ORB
      OUT     T1544 K15
      AND     T1544
      MOV     K50 D1657
      RST     M1750
      RST     M1754
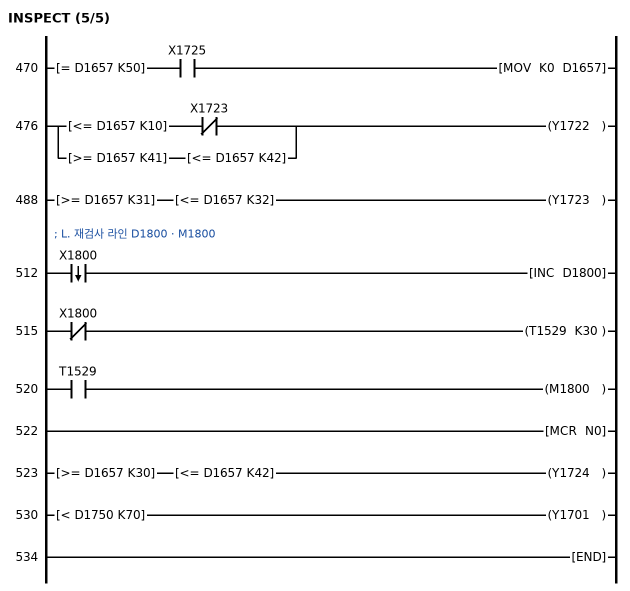
470   LD=     D1657 K50
      AND     X1725
      MOV     K0 D1657
476   LD<=    D1657 K10
      ANI     X1723
      LD>=    D1657 K41
      AND<=   D1657 K42
      ORB
      OUT     Y1722
488   LD>=    D1657 K31
      AND<=   D1657 K32
      OUT     Y1723
; L. 재검사 라인 D1800 · M1800
512   LDF     X1800
      INC     D1800
515   LDI     X1800
      OUT     T1529 K30
520   LD      T1529
      OUT     M1800
522   MCR     N0
523   LD>=    D1657 K30
      AND<=   D1657 K42
      OUT     Y1724
530   LD<     D1750 K70
      OUT     Y1701
534   END
END_PROGRAM

PROGRAM RETEST
